// TIA Portal V21 export
// export: Created 2026-08-21T20:18:53.5001535Z, ExportSetting None, DisplayName Totally Integrated Automation Portal, DisplayVersion V21, DisplayName STEP 7 Professional, DisplayVersion V21, DisplayName STEP 7 Safety, DisplayVersion V21, DisplayName Tech WebApplication, DisplayVersion V21, DisplayName WinCC Basic/Comfort/Advanced, DisplayVersion V21, DisplayName WinCC Professional, DisplayVersion V21, DisplayName WinCC Unified, DisplayVersion V21
FUNCTION "Vlv_Sim" : Void   // FC13, FBD
{ S7_Optimized_Access := 'TRUE' }
// stored: SetENOAutomatically false
BEGIN

REGION Network 1: PT1
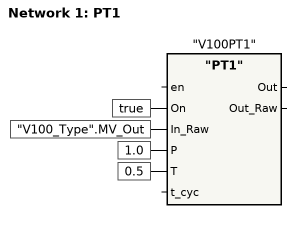
   "V100PT1"(On := true, In_Raw := "V100_Type".MV_Out, P := 1.0, T := 0.5);   // "PT1"
END_REGION
END_FUNCTION
